FUNCTION_BLOCK FB_ForceController
VAR_INPUT
END_VAR
VAR_OUTPUT
END_VAR
VAR
END_VAR

END_FUNCTION_BLOCK

(* stored: Version 1.1.0.1, ProductVersion 3.1.4024.15
   POU FB_ForceController: Id {61d1f3bc-331b-4be7-a710-c3dc213b081e}, SpecialFunc None *)
